(* IEC 61131-3 sources: plc-workbench/experiments/formal_r7/final_recheck/real_model_acknowledge_latch, 2 files *)

(* ---- before.st ---- *)
FUNCTION_BLOCK AcknowledgeLatch
VAR_INPUT
    fault : BOOL;
    acknowledge : BOOL;
END_VAR
VAR_OUTPUT
    alarm : BOOL := FALSE;
END_VAR
VAR
    prevAck : BOOL := FALSE;
    ackRising : BOOL := FALSE;
END_VAR

ackRising := acknowledge AND NOT prevAck;
prevAck := acknowledge;

IF fault THEN
    alarm := TRUE;
ELSIF ackRising THEN
    alarm := FALSE;
END_IF;

END_FUNCTION_BLOCK

(* ---- candidate_final.st ---- *)
FUNCTION_BLOCK AcknowledgeLatch
VAR_INPUT
    fault : BOOL;
    acknowledge : BOOL;
END_VAR
VAR_OUTPUT
    alarm : BOOL := FALSE;
END_VAR
VAR
    prevAck : BOOL := FALSE;
    ackRising : BOOL := FALSE;
END_VAR

ackRising := acknowledge AND NOT prevAck;
prevAck := acknowledge;

IF fault THEN
    alarm := TRUE;
ELSIF ackRising THEN
    alarm := FALSE;
END_IF;

END_FUNCTION_BLOCK
